(* IEC 61131-3 sources: stc/examples/function, 2 files *)

(* ---- function.st ---- *)
FUNCTION F_Sample : INT
  VAR_INPUT
    x : INT;
    y : INT;
  END_VAR
  F_Sample := x + y;
END_FUNCTION;

(* ---- function_no_args.st ---- *)
FUNCTION F_Sample
END_FUNCTION;
